TYPE "DT_REGULATOR_INTERFACE_ALL"
VERSION : 0.1
   STRUCT
      WATER_LEVEL : "DT_REGULATOR_INTERFACE";
      WATER_PRESSURE : "DT_REGULATOR_INTERFACE";
      ACTIVE_POWER : "DT_REGULATOR_INTERFACE";
      OPENNESS : "DT_REGULATOR_INTERFACE";
      SPEED : "DT_REGULATOR_INTERFACE";
      KAPLAN_DISTRIBUTOR : "DT_REGULATOR_INTERFACE";
      KAPLAN_RUNNER : "DT_REGULATOR_INTERFACE";
      FRANCIS_DISTRIBUTOR : "DT_REGULATOR_INTERFACE";
      CROSS_FLOW_VALVE_1 : "DT_REGULATOR_INTERFACE";
      CROSS_FLOW_VALVE_2 : "DT_REGULATOR_INTERFACE";
      PELTON_DEFLECTOR { S7_SetPoint := 'False'} : Array[1..6] of "DT_REGULATOR_INTERFACE";
      PELTON_NOZZLE : Array[1..6] of "DT_REGULATOR_INTERFACE";
      EXC_VOLTAGE : "DT_REGULATOR_INTERFACE";
      EXC_REACTIVE_POWER : "DT_REGULATOR_INTERFACE";
      EXC_POWER_FACTOR : "DT_REGULATOR_INTERFACE";
      Element_25 : "DT_REGULATOR_INTERFACE";
      Element_26 : "DT_REGULATOR_INTERFACE";
      Element_27 : "DT_REGULATOR_INTERFACE";
      Element_28 : "DT_REGULATOR_INTERFACE";
      Element_29 : "DT_REGULATOR_INTERFACE";
      Element_30 : "DT_REGULATOR_INTERFACE";
      Element_31 : "DT_REGULATOR_INTERFACE";
   END_STRUCT;

END_TYPE

